FUNCTION_BLOCK FB_CompI
(*
Function block used to calculate integral typ.

Constructor: 		Patryk Panylo
Company:		E. Riexinger GmbH
Date:			03.06.2014
Version:			1.00

Date:			Revision:		Who:				Comment
dd.mm.yyyy		x.xx			Initials			comment

*)

VAR_INPUT
	(* Enummerations *)

	(* Variables *)
	bEnable								:BOOL := TRUE;					(* Enable FB *)
	lrInSignal								:LREAL;							(* Input signal *)
	lrIntegralValue						:LREAL := 1.0;						(* Integration value in 1/sec *)
	lrTaskCycle							:LREAL := 1.0; 					(* Cycle time *)
	bSetToZero 							:BOOL;							(* Integral set to zero *)
	lrLimitMin								:LREAL := -1E40;					(* Limit minimum *)
	lrLimitMax							:LREAL := 1E40;					(* Limit maximum *)

	(* References *)

	(* Interfaces *)

	(* Instances *)

END_VAR
VAR_OUTPUT
	(* Enummerations *)

	(* Variables *)
	lrOutSignal							:LREAL;							(* Output signal *)
	bLimitMin							:BOOL;							(* Limit minimum reached *)
	bLimitMax							:BOOL;							(* Limit maximum reached *)

	(* References *)

	(* Interfaces *)

	(* Instances *)
END_VAR
VAR
	(* Enummerations *)

	(* Variables *)
	bFirstTime							:BOOL;							(* First cycle *)

	(* References *)

	(* Interfaces *)

	(* Instances *)
	fbIntegral								:FB_Integral;

END_VAR

IF NOT bEnable
THEN

	bLimitMin := FALSE;
	bLimitMax := FALSE;

	fbIntegral(
		bEnable := FALSE,
		lrInSignal := lrInSignal,
		lrIntegralValue := lrIntegralValue,
		lrTaskCycle := lrTaskCycle,
		lrOutSignal := lrOutSignal
	);

	bFirstTime := FALSE;
	RETURN;
END_IF

IF NOT bFirstTime
THEN
	bFirstTime := TRUE;
END_IF

IF bSetToZero
THEN
	lrOutSignal := 0.0;
ELSE

	A_CalcIntegral();

END_IF

A_CheckLimits();

ACTION A_CalcIntegral:

fbIntegral(
	bEnable := TRUE,
	lrInSignal := lrInSignal,
	lrIntegralValue := lrIntegralValue,
	lrTaskCycle := lrTaskCycle,
	lrOutSignal := lrOutSignal
);
END_ACTION

ACTION A_CheckLimits:

(* Check limit the outputs *)
bLimitMin := FALSE;							(* Limit minimum reached *)
bLimitMax := FALSE;							(* Limit maximum reached *)
IF lrOutSignal <= lrLimitMin
THEN
	lrOutSignal := lrLimitMin;
	bLimitMin := TRUE;						(* Limit minimum reached *)

ELSIF  lrOutSignal >= lrLimitMax
THEN
	lrOutSignal := lrLimitMax;
	bLimitMax := TRUE;						(* Limit minimum reached *)

END_IF
END_ACTION

END_FUNCTION_BLOCK

(* stored: Version 1.1.0.1, ProductVersion 3.1.4024.15
   POU FB_CompI: Id {df14b1d2-428d-4320-8d6d-5f46da830245}, SpecialFunc None
   Action A_CalcIntegral: Id {a7b7d660-da6b-4a5e-84bf-1a38f1fd2b3f}
   Action A_CheckLimits: Id {b681348f-c59f-4c72-b4d2-4260be6e505d} *)
